KUKA KRL program: MAIN_1.src

DEF MAIN_1 ( )

;FOLD INI
BAS (#INITMOV,0 )
;ENDFOLD (INI)

;FOLD STARTPOS
$BWDSTART = FALSE
PDAT_ACT = PDEFAULT
BAS(#PTP_DAT)
FDAT_ACT = {TOOL_NO 0,BASE_NO 0,IPO_FRAME #BASE}
BAS(#FRAMES)
;ENDFOLD

;FOLD SET DEFAULT SPEED
$VEL.CP=0.2
BAS(#VEL_PTP,100)
BAS(#TOOL,0)
BAS(#BASE,0)
;ENDFOLD

PTP $AXIS_ACT ; skip BCO quickly

$ACC.CP = 2.00000
; Program generated by RoboDK v5.6.9 for RoboDK Industrial on 26/02/2024 09:58:20
; Using nominal kinematics.
PTP {A1 -0.00000,A2 0.00000,A3 0.00000,A4 0.00000,A5 0.00000,A6 -0.00000}
PTP {A1 0.00000,A2 3.21124,A3 -15.42370,A4 0.00000,A5 12.21250,A6 -0.00000}
CR_PROCESS_FILE("MAIN_1.csv", 1, -1, "OK" )
$OUT[5]=TRUE
$OUT[5]=TRUE
$OUT[5]=0.5
$OUT[5]=true
$ANOUT[5]=TRUE
$ANOUT[5]=TRUE
$ANOUT[5]=0.5
$ANOUT[5]=true
var=val
var=val
WAIT FOR ($IN[5]==TRUE)
WAIT FOR ($IN[5]==TRUE)
WAIT FOR ($IN[5]==0.5)
WAIT FOR ($IN[5]==true)
START_TIMER:
$TIMER_STOP[1]=TRUE
$TIMER_FLAG[1]=FALSE
$TIMER[1]=0.100
$TIMER_STOP[1]=FALSE
WAIT FOR ($IN[5]==TRUE OR $TIMER_FLAG[1])
$TIMER_STOP[1]=TRUE
IF $TIMER_FLAG[1]== TRUE THEN
    HALT ; Timed out!
    GOTO START_TIMER
ENDIF
WAIT FOR (var==val)
START_TIMER:
$TIMER_STOP[1]=TRUE
$TIMER_FLAG[1]=FALSE
$TIMER[1]=0.100
$TIMER_STOP[1]=FALSE
WAIT FOR (var==val OR $TIMER_FLAG[1])
$TIMER_STOP[1]=TRUE
IF $TIMER_FLAG[1]== TRUE THEN
    HALT ; Timed out!
    GOTO START_TIMER
ENDIF
; Insert Comment
$APO.CPTP = 10
$APO.CDIS = 10.000
PTP {A1 -29.33220,A2 46.67700,A3 -0.02452,A4 26.54560,A5 25.39570,A6 -51.63400} C_PTP
$OUT[5]=TRUE
$APO.CPTP = 10
$APO.CDIS = 10.000
; Linear movement using joint targets is not supported. Change the target type to cartesian or use a joint movement.
; MoveSearch command not implemented
$OUT[5]=FALSE
$APO.CPTP = 10
$APO.CDIS = 10.000
$APO.CPTP = 25
$APO.CDIS = 25.000
PTP {A1 52.18600,A2 45.67580,A3 6.92000,A4 66.73420,A5 19.93230,A6 -92.73000} C_PTP
PTP {A1 -0.00000,A2 0.00000,A3 0.00000,A4 0.00000,A5 0.00000,A6 -0.00000}
PTP {A1 88.67600,A2 29.60160,A3 -6.42883,A4 -1.98422,A5 49.47920,A6 4.54769}
PTP {A1 -0.00000,A2 0.00000,A3 0.00000,A4 0.00000,A5 0.00000,A6 -0.00000}
$APO.CPTP = 1
$APO.CDIS = 1.000
; Show Tool 1
PTP {A1 -68.09030,A2 24.20190,A3 26.78550,A4 38.21340,A5 36.20170,A6 -98.79640} C_PTP
PTP {A1 -29.33220,A2 46.67700,A3 -0.02452,A4 26.54560,A5 25.39570,A6 -51.63400} C_PTP
WAIT FOR ($IN[1]==TRUE)
END
